// TIA Portal V19 export
VAR_GLOBAL   // PLC tag table "Press"
   DI_NCP45_Press AT %I8.3 : Bool;
   "DI_Press_ReadyCycleComplete/Power" AT %I13.0 : Bool;
   "DI_Press_TopPosition/emg_Stop" AT %I13.1 : Bool;
   "DI_AirPressure_OK/Ready" AT %I13.2 : Bool;
   "DI_Motor_Running/MainMotor" AT %I13.3 : Bool;
   DI_MotorOverload AT %I13.4 : Bool;
   DI_Disconector_ON AT %I13.5 : Bool;
   "DI_Left/Right TrayStuck" AT %I13.6 : Bool;
   "DQ_Press_Run/Operate" AT %Q17.0 : Bool;
   DQ_Press_Reset AT %Q17.1 : Bool;
   "DQ_Press_FWD/MotorsStart" AT %Q17.2 : Bool;
   "DQ_Press_REV/MotorStop" AT %Q17.3 : Bool;
   "DQ_Press_Jog/Power" AT %Q17.4 : Bool;
   "DQ_Press_Cycle_Mode/Stroke" AT %Q17.5 : Bool;
   DQ_Press_Air AT %Q17.6 : Bool;
END_VAR
